Yaskawa INFORM job: CALIBPOSON.JBI

/JOB
//NAME CALIBPOSON
///FOLDERNAME FOLDER003
//POS
///NPOS 0,0,0,0,0,0
//INST
///DATE 2021/11/07 16:16
///ATTR SC,RW
///GROUP1 RB1
NOP
SET B010 1
TIMER T=2.00
WAIT B010=0
END
